(* IEC 61131-3 sources: plc-st-coding-agent/progress/evidence/f14_v6_public_pilot_20261112/jobs/custom_deepseek-v4pro (part 2) *)

(* ---- public-medium-04.candidate_01.st ---- *)
FUNCTION_BLOCK FB_TemperatureControl
VAR_INPUT
    TemperatureSensorInput : REAL;
    SetTemperature : REAL;
END_VAR
VAR_OUTPUT
    CurrentTemperature : REAL;
    SetTempDisplay : REAL;
    HeaterStatus : BOOL;
    OverheatProtection : BOOL;
    HeaterOutput : BOOL;
END_VAR
VAR
    sensor_fault : BOOL;
    heater_request : BOOL;
    heater_timer_in : BOOL;
    overheat_active : BOOL;
    HeatingTimer : TON;
    CoolingTimer : TON;
END_VAR

(* ENGINEERING_CONTRACT
   O1 CurrentTemperature: always copies TemperatureSensorInput; no fault suppression; units = input units (PUB006/PUB007).
   O2 SetTempDisplay: always copies SetTemperature; units same as input (PUB006/PUB007).
   O3 HeaterStatus: copies final HeaterOutput; true while actual heater command active (PUB006/PUB007).
   O4 OverheatProtection: latched TRUE when HeatingTimer reaches T#5S; holds TRUE while CoolingTimer < T#3S; auto-clears after T#3S; no external reset (PUB005/PUB006).
   O5 HeaterOutput: TRUE when sensor input in [0,100] and TemperatureSensorInput < SetTemperature and not overheat-active; FALSE on sensor fault, overheat, or temp >= set (PUB003/PUB004/PUB005/PUB008).
   State retention: OverheatProtection retained during 3s wait; HeatingTimer resets whenever HeaterOutput is false; CoolingTimer resets when overheat inactive.
   Same-scan priority: overheat set and HeaterOutput forced FALSE in same timer-trigger scan; when cooling timer completes, HeaterOutput may turn on same scan if setpoint condition still true.
   Boundaries: strict < for low-temperature start; fault uses <0.0 or >100.0; exact 0/100 valid; T#5S and T#3S are TIME constants.
*)
(* CONTRACT_RULES [] *)

sensor_fault := (TemperatureSensorInput < 0.0) OR (TemperatureSensorInput > 100.0);
heater_request := (NOT sensor_fault) AND (TemperatureSensorInput < SetTemperature);

IF overheat_active THEN
    heater_timer_in := FALSE;
ELSE
    heater_timer_in := heater_request;
END_IF;

HeatingTimer(IN := heater_timer_in, PT := T#5S);
IF HeatingTimer.Q THEN
    overheat_active := TRUE;
    heater_timer_in := FALSE;
END_IF;

CoolingTimer(IN := overheat_active, PT := T#3S);
IF overheat_active AND CoolingTimer.Q THEN
    overheat_active := FALSE;
END_IF;

HeaterOutput := heater_request AND NOT overheat_active;
CurrentTemperature := TemperatureSensorInput;
SetTempDisplay := SetTemperature;
HeaterStatus := HeaterOutput;
OverheatProtection := overheat_active;

END_FUNCTION_BLOCK

(* ---- public-medium-04.candidate_02.st ---- *)
FUNCTION_BLOCK FB_TemperatureControl
VAR_INPUT
    TemperatureSensorInput : REAL;
    SetTemperature : REAL;
END_VAR
VAR_OUTPUT
    CurrentTemperature : REAL;
    SetTempDisplay : REAL;
    HeaterStatus : BOOL;
    OverheatProtection : BOOL;
    HeaterOutput : BOOL;
END_VAR
VAR
    sensor_fault : BOOL;
    heater_request : BOOL;
    overheat_active : BOOL;
    tmp_heater_in : BOOL;
    HeatingTimer : TON;
    CoolingTimer : TON;
END_VAR

(* ENGINEERING_CONTRACT
   O1 CurrentTemperature: always copies TemperatureSensorInput; no fault suppression; units = input units (PUB006/PUB007).
   O2 SetTempDisplay: always copies SetTemperature; units same as input (PUB006/PUB007).
   O3 HeaterStatus: copies final HeaterOutput; true while actual heater command active (PUB006/PUB007).
   O4 OverheatProtection: latched TRUE when HeatingTimer reaches T#5S; holds TRUE while CoolingTimer < T#3S; auto-clears after T#3S; no external reset (PUB005/PUB006).
   O5 HeaterOutput: TRUE when sensor input in [0,100] and TemperatureSensorInput < SetTemperature and not overheat-active; FALSE on sensor fault, overheat, or temp >= set (PUB003/PUB004/PUB005/PUB008).
   State retention: OverheatProtection retained during 3s wait; HeatingTimer resets whenever HeaterOutput is false; CoolingTimer resets when overheat inactive.
   Same-scan priority: overheat set and HeaterOutput forced FALSE in same timer-trigger scan; when cooling timer completes, HeaterOutput may turn on same scan if setpoint condition still true.
   Boundaries: strict < for low-temperature start; fault uses <0.0 or >100.0; exact 0/100 valid; T#5S and T#3S are TIME constants.
*)
(* CONTRACT_RULES [] *)

sensor_fault := (TemperatureSensorInput < 0.0) OR (TemperatureSensorInput > 100.0);
heater_request := (NOT sensor_fault) AND (TemperatureSensorInput < SetTemperature);

(* Desired heating timer enable before possible cooling-timer completion. *)
tmp_heater_in := heater_request AND NOT overheat_active;

(* First HeatingTimer call: handle normal heating and detect overheat trigger. *)
HeatingTimer(IN := tmp_heater_in, PT := T#5S);
IF HeatingTimer.Q THEN
    overheat_active := TRUE;
    tmp_heater_in := FALSE;
END_IF;

(* CoolingTimer call: starts if overheat just triggered, clears after 3 s. *)
CoolingTimer(IN := overheat_active, PT := T#3S);
IF overheat_active AND CoolingTimer.Q THEN
    overheat_active := FALSE;
END_IF;

HeaterOutput := heater_request AND NOT overheat_active;

(* Ensure HeatingTimer starts immediately when heater turns on in this scan.
   Also reset immediately when heater turns off to avoid one-scan timer drift. *)
IF HeaterOutput AND NOT tmp_heater_in THEN
    HeatingTimer(IN := TRUE, PT := T#5S);
ELSIF (NOT HeaterOutput) AND tmp_heater_in THEN
    HeatingTimer(IN := FALSE, PT := T#5S);
END_IF;

CurrentTemperature := TemperatureSensorInput;
SetTempDisplay := SetTemperature;
HeaterStatus := HeaterOutput;
OverheatProtection := overheat_active;

END_FUNCTION_BLOCK

(* ---- public-medium-04.candidate_03.st ---- *)
FUNCTION_BLOCK FB_TemperatureControl
VAR_INPUT
    TemperatureSensorInput : REAL;
    SetTemperature : REAL;
END_VAR
VAR_OUTPUT
    CurrentTemperature : REAL;
    SetTempDisplay : REAL;
    HeaterStatus : BOOL;
    OverheatProtection : BOOL;
    HeaterOutput : BOOL;
END_VAR
VAR
    sensor_fault : BOOL;
    heater_request : BOOL;
    overheat_active : BOOL;
    tmp_heater_in : BOOL;
    HeatingTimer : TON;
    CoolingTimer : TON;
END_VAR

(* ENGINEERING_CONTRACT
   O1 CurrentTemperature: always copies TemperatureSensorInput; no fault suppression; units = input units (PUB006/PUB007).
   O2 SetTempDisplay: always copies SetTemperature; units same as input (PUB006/PUB007).
   O3 HeaterStatus: copies final HeaterOutput; true while actual heater command active (PUB006/PUB007).
   O4 OverheatProtection: latched TRUE when HeatingTimer reaches T#5S; holds TRUE while CoolingTimer < T#3S; auto-clears after T#3S; no external reset (PUB005/PUB006).
   O5 HeaterOutput: TRUE when sensor input in [0,100] and TemperatureSensorInput < SetTemperature and not overheat-active; FALSE on sensor fault, overheat, or temp >= set (PUB003/PUB004/PUB005/PUB008).
   State retention: OverheatProtection retained during 3s wait; HeatingTimer resets whenever HeaterOutput is false; CoolingTimer resets when overheat inactive.
   Same-scan priority: overheat set and HeaterOutput forced FALSE in same timer-trigger scan; when cooling timer completes, HeaterOutput may turn on same scan if setpoint condition still true.
   Boundaries: strict < for low-temperature start; fault uses <0.0 or >100.0; exact 0/100 valid; T#5S and T#3S are TIME constants.
*)
(* CONTRACT_RULES [] *)

sensor_fault := (TemperatureSensorInput < 0.0) OR (TemperatureSensorInput > 100.0);
heater_request := (NOT sensor_fault) AND (TemperatureSensorInput < SetTemperature);

(* Single HeatingTimer call with enable = heater_request AND NOT overheat_active. *)
tmp_heater_in := heater_request AND NOT overheat_active;
HeatingTimer(IN := tmp_heater_in, PT := T#5S);

IF HeatingTimer.Q THEN
    overheat_active := TRUE;
END_IF;

(* Single CoolingTimer call with enable = overheat_active. *)
CoolingTimer(IN := overheat_active, PT := T#3S);
IF CoolingTimer.Q THEN
    overheat_active := FALSE;
END_IF;

HeaterOutput := heater_request AND NOT overheat_active;

CurrentTemperature := TemperatureSensorInput;
SetTempDisplay := SetTemperature;
HeaterStatus := HeaterOutput;
OverheatProtection := overheat_active;

END_FUNCTION_BLOCK

(* ---- public-medium-04.candidate_04.st ---- *)
FUNCTION_BLOCK FB_TemperatureControl
VAR_INPUT
    TemperatureSensorInput : REAL;
    SetTemperature : REAL;
END_VAR
VAR_OUTPUT
    CurrentTemperature : REAL;
    SetTempDisplay : REAL;
    HeaterStatus : BOOL;
    OverheatProtection : BOOL;
    HeaterOutput : BOOL;
END_VAR
VAR
    sensor_fault : BOOL;
    heater_request : BOOL;
    overheat_active : BOOL;
    HeatingTimer : TON;
    CoolingTimer : TON;
END_VAR

(* ENGINEERING_CONTRACT
   O1 CurrentTemperature: always copies TemperatureSensorInput; no fault suppression; units = input units (PUB006/PUB007).
   O2 SetTempDisplay: always copies SetTemperature; units same as input (PUB006/PUB007).
   O3 HeaterStatus: copies final HeaterOutput; true while actual heater command active (PUB006/PUB007).
   O4 OverheatProtection: latched TRUE when HeatingTimer reaches T#5S; holds TRUE while CoolingTimer < T#3S; auto-clears after T#3S; no external reset (PUB005/PUB006).
   O5 HeaterOutput: TRUE when sensor input in [0,100] and TemperatureSensorInput < SetTemperature and not overheat-active; FALSE on sensor fault, overheat, or temp >= set (PUB003/PUB004/PUB005/PUB008).
   State retention: OverheatProtection retained during 3s wait; HeatingTimer resets whenever HeaterOutput is false; CoolingTimer resets when overheat inactive.
   Same-scan priority: overheat set and HeaterOutput forced FALSE in same timer-trigger scan; when cooling timer completes, HeaterOutput may turn on same scan if setpoint condition still true.
   Boundaries: strict < for low-temperature start; fault uses <0.0 or >100.0; exact 0/100 valid; T#5S and T#3S are TIME constants.
*)
(* CONTRACT_RULES [] *)

sensor_fault := (TemperatureSensorInput < 0.0) OR (TemperatureSensorInput > 100.0);
heater_request := (NOT sensor_fault) AND (TemperatureSensorInput < SetTemperature);

(* Initial heater output based on current overheat state *)
HeaterOutput := heater_request AND NOT overheat_active;

(* Heating timer: active only when heater is actually on *)
HeatingTimer(IN := HeaterOutput, PT := T#5S);
IF HeatingTimer.Q THEN
    overheat_active := TRUE;
    HeaterOutput := FALSE;   (* force off immediately *)
    HeatingTimer(IN := FALSE, PT := T#5S); (* reset timer *)
END_IF;

(* Cooling timer: active while overheat protection is latched *)
CoolingTimer(IN := overheat_active, PT := T#3S);
IF overheat_active AND CoolingTimer.Q THEN
    overheat_active := FALSE;
    HeaterOutput := heater_request; (* may turn on again if still low *)
    CoolingTimer(IN := FALSE, PT := T#3S); (* reset cooling timer *)
END_IF;

CurrentTemperature := TemperatureSensorInput;
SetTempDisplay := SetTemperature;
HeaterStatus := HeaterOutput;
OverheatProtection := overheat_active;

END_FUNCTION_BLOCK

(* ---- public-medium-04.raw_candidate_01.st ---- *)
FUNCTION_BLOCK FB_TemperatureControl
VAR_INPUT
    TemperatureSensorInput : REAL;
    SetTemperature : REAL;
END_VAR
VAR_OUTPUT
    CurrentTemperature : REAL;
    SetTempDisplay : REAL;
    HeaterStatus : BOOL;
    OverheatProtection : BOOL;
    HeaterOutput : BOOL;
END_VAR
VAR
    sensor_fault : BOOL;
    heater_request : BOOL;
    heater_timer_in : BOOL;
    overheat_active : BOOL;
    HeatingTimer : TON;
    CoolingTimer : TON;
END_VAR

(* ENGINEERING_CONTRACT
   O1 CurrentTemperature: always copies TemperatureSensorInput; no fault suppression; units = input units (PUB006/PUB007).
   O2 SetTempDisplay: always copies SetTemperature; units same as input (PUB006/PUB007).
   O3 HeaterStatus: copies final HeaterOutput; true while actual heater command active (PUB006/PUB007).
   O4 OverheatProtection: latched TRUE when HeatingTimer reaches T#5S; holds TRUE while CoolingTimer < T#3S; auto-clears after T#3S; no external reset (PUB005/PUB006).
   O5 HeaterOutput: TRUE when sensor input in [0,100] and TemperatureSensorInput < SetTemperature and not overheat-active; FALSE on sensor fault, overheat, or temp >= set (PUB003/PUB004/PUB005/PUB008).
   State retention: OverheatProtection retained during 3s wait; HeatingTimer resets whenever HeaterOutput is false; CoolingTimer resets when overheat inactive.
   Same-scan priority: overheat set and HeaterOutput forced FALSE in same timer-trigger scan; when cooling timer completes, HeaterOutput may turn on same scan if setpoint condition still true.
   Boundaries: strict < for low-temperature start; fault uses <0.0 or >100.0; exact 0/100 valid; T#5S and T#3S are TIME constants.
*)
(* CONTRACT_RULES [] *)

sensor_fault := (TemperatureSensorInput < 0.0) OR (TemperatureSensorInput > 100.0);
heater_request := (NOT sensor_fault) AND (TemperatureSensorInput < SetTemperature);

IF overheat_active THEN
    heater_timer_in := FALSE;
ELSE
    heater_timer_in := heater_request;
END_IF;

HeatingTimer(IN := heater_timer_in, PT := T#5S);
IF HeatingTimer.Q THEN
    overheat_active := TRUE;
    heater_timer_in := FALSE;
END_IF;

CoolingTimer(IN := overheat_active, PT := T#3S);
IF overheat_active AND CoolingTimer.Q THEN
    overheat_active := FALSE;
END_IF;

HeaterOutput := heater_request AND NOT overheat_active;
CurrentTemperature := TemperatureSensorInput;
SetTempDisplay := SetTemperature;
HeaterStatus := HeaterOutput;
OverheatProtection := overheat_active;

END_FUNCTION_BLOCK

(* ---- public-medium-04.raw_candidate_02.st ---- *)
FUNCTION_BLOCK FB_TemperatureControl
VAR_INPUT
    TemperatureSensorInput : REAL;
    SetTemperature : REAL;
END_VAR
VAR_OUTPUT
    CurrentTemperature : REAL;
    SetTempDisplay : REAL;
    HeaterStatus : BOOL;
    OverheatProtection : BOOL;
    HeaterOutput : BOOL;
END_VAR
VAR
    sensor_fault : BOOL;
    heater_request : BOOL;
    overheat_active : BOOL;
    tmp_heater_in : BOOL;
    HeatingTimer : TON;
    CoolingTimer : TON;
END_VAR

(* ENGINEERING_CONTRACT
   O1 CurrentTemperature: always copies TemperatureSensorInput; no fault suppression; units = input units (PUB006/PUB007).
   O2 SetTempDisplay: always copies SetTemperature; units same as input (PUB006/PUB007).
   O3 HeaterStatus: copies final HeaterOutput; true while actual heater command active (PUB006/PUB007).
   O4 OverheatProtection: latched TRUE when HeatingTimer reaches T#5S; holds TRUE while CoolingTimer < T#3S; auto-clears after T#3S; no external reset (PUB005/PUB006).
   O5 HeaterOutput: TRUE when sensor input in [0,100] and TemperatureSensorInput < SetTemperature and not overheat-active; FALSE on sensor fault, overheat, or temp >= set (PUB003/PUB004/PUB005/PUB008).
   State retention: OverheatProtection retained during 3s wait; HeatingTimer resets whenever HeaterOutput is false; CoolingTimer resets when overheat inactive.
   Same-scan priority: overheat set and HeaterOutput forced FALSE in same timer-trigger scan; when cooling timer completes, HeaterOutput may turn on same scan if setpoint condition still true.
   Boundaries: strict < for low-temperature start; fault uses <0.0 or >100.0; exact 0/100 valid; T#5S and T#3S are TIME constants.
*)
(* CONTRACT_RULES [] *)

sensor_fault := (TemperatureSensorInput < 0.0) OR (TemperatureSensorInput > 100.0);
heater_request := (NOT sensor_fault) AND (TemperatureSensorInput < SetTemperature);

(* Desired heating timer enable before possible cooling-timer completion. *)
tmp_heater_in := heater_request AND NOT overheat_active;

(* First HeatingTimer call: handle normal heating and detect overheat trigger. *)
HeatingTimer(IN := tmp_heater_in, PT := T#5S);
IF HeatingTimer.Q THEN
    overheat_active := TRUE;
    tmp_heater_in := FALSE;
END_IF;

(* CoolingTimer call: starts if overheat just triggered, clears after 3 s. *)
CoolingTimer(IN := overheat_active, PT := T#3S);
IF overheat_active AND CoolingTimer.Q THEN
    overheat_active := FALSE;
END_IF;

HeaterOutput := heater_request AND NOT overheat_active;

(* Ensure HeatingTimer starts immediately when heater turns on in this scan.
   Also reset immediately when heater turns off to avoid one-scan timer drift. *)
IF HeaterOutput AND NOT tmp_heater_in THEN
    HeatingTimer(IN := TRUE, PT := T#5S);
ELSIF (NOT HeaterOutput) AND tmp_heater_in THEN
    HeatingTimer(IN := FALSE, PT := T#5S);
END_IF;

CurrentTemperature := TemperatureSensorInput;
SetTempDisplay := SetTemperature;
HeaterStatus := HeaterOutput;
OverheatProtection := overheat_active;

END_FUNCTION_BLOCK

(* ---- public-medium-04.raw_candidate_03.st ---- *)
FUNCTION_BLOCK FB_TemperatureControl
VAR_INPUT
    TemperatureSensorInput : REAL;
    SetTemperature : REAL;
END_VAR
VAR_OUTPUT
    CurrentTemperature : REAL;
    SetTempDisplay : REAL;
    HeaterStatus : BOOL;
    OverheatProtection : BOOL;
    HeaterOutput : BOOL;
END_VAR
VAR
    sensor_fault : BOOL;
    heater_request : BOOL;
    overheat_active : BOOL;
    tmp_heater_in : BOOL;
    HeatingTimer : TON;
    CoolingTimer : TON;
END_VAR

(* ENGINEERING_CONTRACT
   O1 CurrentTemperature: always copies TemperatureSensorInput; no fault suppression; units = input units (PUB006/PUB007).
   O2 SetTempDisplay: always copies SetTemperature; units same as input (PUB006/PUB007).
   O3 HeaterStatus: copies final HeaterOutput; true while actual heater command active (PUB006/PUB007).
   O4 OverheatProtection: latched TRUE when HeatingTimer reaches T#5S; holds TRUE while CoolingTimer < T#3S; auto-clears after T#3S; no external reset (PUB005/PUB006).
   O5 HeaterOutput: TRUE when sensor input in [0,100] and TemperatureSensorInput < SetTemperature and not overheat-active; FALSE on sensor fault, overheat, or temp >= set (PUB003/PUB004/PUB005/PUB008).
   State retention: OverheatProtection retained during 3s wait; HeatingTimer resets whenever HeaterOutput is false; CoolingTimer resets when overheat inactive.
   Same-scan priority: overheat set and HeaterOutput forced FALSE in same timer-trigger scan; when cooling timer completes, HeaterOutput may turn on same scan if setpoint condition still true.
   Boundaries: strict < for low-temperature start; fault uses <0.0 or >100.0; exact 0/100 valid; T#5S and T#3S are TIME constants.
*)
(* CONTRACT_RULES [] *)

sensor_fault := (TemperatureSensorInput < 0.0) OR (TemperatureSensorInput > 100.0);
heater_request := (NOT sensor_fault) AND (TemperatureSensorInput < SetTemperature);

(* Single HeatingTimer call with enable = heater_request AND NOT overheat_active. *)
tmp_heater_in := heater_request AND NOT overheat_active;
HeatingTimer(IN := tmp_heater_in, PT := T#5S);

IF HeatingTimer.Q THEN
    overheat_active := TRUE;
END_IF;

(* Single CoolingTimer call with enable = overheat_active. *)
CoolingTimer(IN := overheat_active, PT := T#3S);
IF CoolingTimer.Q THEN
    overheat_active := FALSE;
END_IF;

HeaterOutput := heater_request AND NOT overheat_active;

CurrentTemperature := TemperatureSensorInput;
SetTempDisplay := SetTemperature;
HeaterStatus := HeaterOutput;
OverheatProtection := overheat_active;

END_FUNCTION_BLOCK

(* ---- public-medium-04.raw_candidate_04.st ---- *)
FUNCTION_BLOCK FB_TemperatureControl
VAR_INPUT
    TemperatureSensorInput : REAL;
    SetTemperature : REAL;
END_VAR
VAR_OUTPUT
    CurrentTemperature : REAL;
    SetTempDisplay : REAL;
    HeaterStatus : BOOL;
    OverheatProtection : BOOL;
    HeaterOutput : BOOL;
END_VAR
VAR
    sensor_fault : BOOL;
    heater_request : BOOL;
    overheat_active : BOOL;
    HeatingTimer : TON;
    CoolingTimer : TON;
END_VAR

(* ENGINEERING_CONTRACT
   O1 CurrentTemperature: always copies TemperatureSensorInput; no fault suppression; units = input units (PUB006/PUB007).
   O2 SetTempDisplay: always copies SetTemperature; units same as input (PUB006/PUB007).
   O3 HeaterStatus: copies final HeaterOutput; true while actual heater command active (PUB006/PUB007).
   O4 OverheatProtection: latched TRUE when HeatingTimer reaches T#5S; holds TRUE while CoolingTimer < T#3S; auto-clears after T#3S; no external reset (PUB005/PUB006).
   O5 HeaterOutput: TRUE when sensor input in [0,100] and TemperatureSensorInput < SetTemperature and not overheat-active; FALSE on sensor fault, overheat, or temp >= set (PUB003/PUB004/PUB005/PUB008).
   State retention: OverheatProtection retained during 3s wait; HeatingTimer resets whenever HeaterOutput is false; CoolingTimer resets when overheat inactive.
   Same-scan priority: overheat set and HeaterOutput forced FALSE in same timer-trigger scan; when cooling timer completes, HeaterOutput may turn on same scan if setpoint condition still true.
   Boundaries: strict < for low-temperature start; fault uses <0.0 or >100.0; exact 0/100 valid; T#5S and T#3S are TIME constants.
*)
(* CONTRACT_RULES [] *)

sensor_fault := (TemperatureSensorInput < 0.0) OR (TemperatureSensorInput > 100.0);
heater_request := (NOT sensor_fault) AND (TemperatureSensorInput < SetTemperature);

(* Initial heater output based on current overheat state *)
HeaterOutput := heater_request AND NOT overheat_active;

(* Heating timer: active only when heater is actually on *)
HeatingTimer(IN := HeaterOutput, PT := T#5S);
IF HeatingTimer.Q THEN
    overheat_active := TRUE;
    HeaterOutput := FALSE;   (* force off immediately *)
    HeatingTimer(IN := FALSE, PT := T#5S); (* reset timer *)
END_IF;

(* Cooling timer: active while overheat protection is latched *)
CoolingTimer(IN := overheat_active, PT := T#3S);
IF overheat_active AND CoolingTimer.Q THEN
    overheat_active := FALSE;
    HeaterOutput := heater_request; (* may turn on again if still low *)
    CoolingTimer(IN := FALSE, PT := T#3S); (* reset cooling timer *)
END_IF;

CurrentTemperature := TemperatureSensorInput;
SetTempDisplay := SetTemperature;
HeaterStatus := HeaterOutput;
OverheatProtection := overheat_active;

END_FUNCTION_BLOCK

(* ---- public-medium-08.candidate_01.st ---- *)
(* ENGINEERING_CONTRACT
 * Output ipValue: computed each scan (PUB001/PUB003); no retention.
 * Reset/deactivation: ipValue := 0 for malformed, nondigit, wrong segment count, or range error (PUB004).
 * Same-scan priority: only ipText drives ipValue; no competing commands or latches.
 * Units/boundaries: each decimal segment 0..255 (PUB002); assembled network byte order into UDINT (PUB003).
 * Valid 0.0.0.0 yields UDINT 0, indistinguishable from invalid by value only.
 * Leading zeros are accepted; PUB002 defines value range and nonempty digits, no max length.
 * String indexing is zero-based BYTE; ASCII digits 48..57 and dot 46 are the only accepted characters.
 *)

(* CONTRACT_RULES [] *)

FUNCTION_BLOCK FB_IPv4Parser
VAR_INPUT
    ipText : STRING(254);
END_VAR
VAR_OUTPUT
    ipValue : UDINT;
END_VAR
VAR
    local_i : INT;
    local_len : INT;
    local_code : INT;
    local_digit_count : INT;
    local_dot_count : INT;
    local_segment_value : UDINT;
    local_segment_invalid : BOOL;
    local_valid : BOOL;
    local_segments : ARRAY[0..3] OF UDINT;
END_VAR

ipValue := 0;
local_valid := TRUE;
local_len := LEN(ipText);
local_digit_count := 0;
local_dot_count := 0;
local_segment_value := 0;
local_segment_invalid := FALSE;
local_segments[0] := 0;
local_segments[1] := 0;
local_segments[2] := 0;
local_segments[3] := 0;

IF local_len = 0 THEN
    local_valid := FALSE;
END_IF;

FOR local_i := 0 TO local_len - 1 DO
    local_code := BYTE_TO_INT(ipText[local_i]);

    IF (local_code >= 48) AND (local_code <= 57) THEN
        local_digit_count := local_digit_count + 1;
        IF NOT local_segment_invalid THEN
            local_segment_value := local_segment_value * UDINT#10 + INT_TO_UDINT(local_code - 48);
            IF local_segment_value > UDINT#255 THEN
                local_segment_invalid := TRUE;
                local_valid := FALSE;
            END_IF;
        END_IF;

    ELSIF local_code = 46 THEN
        IF (local_digit_count = 0) OR local_segment_invalid OR (local_dot_count >= 3) THEN
            local_valid := FALSE;
        ELSE
            local_segments[local_dot_count] := local_segment_value;
        END_IF;

        local_dot_count := local_dot_count + 1;
        local_digit_count := 0;
        local_segment_value := 0;
        local_segment_invalid := FALSE;

    ELSE
        local_valid := FALSE;
    END_IF;
END_FOR;

IF local_valid AND (local_digit_count > 0) AND (NOT local_segment_invalid) AND (local_dot_count = 3) THEN
    local_segments[3] := local_segment_value;
    ipValue := SHL(local_segments[0], 24)
               OR SHL(local_segments[1], 16)
               OR SHL(local_segments[2], 8)
               OR local_segments[3];
ELSE
    ipValue := 0;
END_IF;

END_FUNCTION_BLOCK

(* ---- public-medium-08.raw_candidate_01.st ---- *)
(* ENGINEERING_CONTRACT
 * Output ipValue: computed each scan (PUB001/PUB003); no retention.
 * Reset/deactivation: ipValue := 0 for malformed, nondigit, wrong segment count, or range error (PUB004).
 * Same-scan priority: only ipText drives ipValue; no competing commands or latches.
 * Units/boundaries: each decimal segment 0..255 (PUB002); assembled network byte order into UDINT (PUB003).
 * Valid 0.0.0.0 yields UDINT 0, indistinguishable from invalid by value only.
 * Leading zeros are accepted; PUB002 defines value range and nonempty digits, no max length.
 * String indexing is zero-based BYTE; ASCII digits 48..57 and dot 46 are the only accepted characters.
 *)

(* CONTRACT_RULES [] *)

FUNCTION_BLOCK FB_IPv4Parser
VAR_INPUT
    ipText : STRING(254);
END_VAR
VAR_OUTPUT
    ipValue : UDINT;
END_VAR
VAR
    local_i : INT;
    local_len : INT;
    local_code : INT;
    local_digit_count : INT;
    local_dot_count : INT;
    local_segment_value : UDINT;
    local_segment_invalid : BOOL;
    local_valid : BOOL;
    local_segments : ARRAY[0..3] OF UDINT;
END_VAR

ipValue := 0;
local_valid := TRUE;
local_len := LEN(ipText);
local_digit_count := 0;
local_dot_count := 0;
local_segment_value := 0;
local_segment_invalid := FALSE;
local_segments[0] := 0;
local_segments[1] := 0;
local_segments[2] := 0;
local_segments[3] := 0;

IF local_len = 0 THEN
    local_valid := FALSE;
END_IF;

FOR local_i := 0 TO local_len - 1 DO
    local_code := BYTE_TO_INT(ipText[local_i]);

    IF (local_code >= 48) AND (local_code <= 57) THEN
        local_digit_count := local_digit_count + 1;
        IF NOT local_segment_invalid THEN
            local_segment_value := local_segment_value * UDINT#10 + INT_TO_UDINT(local_code - 48);
            IF local_segment_value > UDINT#255 THEN
                local_segment_invalid := TRUE;
                local_valid := FALSE;
            END_IF;
        END_IF;

    ELSIF local_code = 46 THEN
        IF (local_digit_count = 0) OR local_segment_invalid OR (local_dot_count >= 3) THEN
            local_valid := FALSE;
        ELSE
            local_segments[local_dot_count] := local_segment_value;
        END_IF;

        local_dot_count := local_dot_count + 1;
        local_digit_count := 0;
        local_segment_value := 0;
        local_segment_invalid := FALSE;

    ELSE
        local_valid := FALSE;
    END_IF;
END_FOR;

IF local_valid AND (local_digit_count > 0) AND (NOT local_segment_invalid) AND (local_dot_count = 3) THEN
    local_segments[3] := local_segment_value;
    ipValue := SHL(local_segments[0], 24)
               OR SHL(local_segments[1], 16)
               OR SHL(local_segments[2], 8)
               OR local_segments[3];
ELSE
    ipValue := 0;
END_IF;

END_FUNCTION_BLOCK
